Fanuc KAREL source: KO00124.KL

PROGRAM KO00124
%NOLOCKGROUP
VAR
  A: ARRAY[2] OF SHORT
  B: REAL
  OUT: REAL
BEGIN
  A[1] = 1
  B = 2
  OUT = ATAN2(A[1], B)
END KO00124
